TYPE ST_PolarIIChamber_HolderRotateServiceCtrl :
STRUCT
	OPR : ST_ServiceCtrl;
	MoveVelocityCW : ST_ServiceCtrl;
	MoveVelocityCCW : ST_ServiceCtrl;
	MoveModulo : ST_ServiceCtrl;
END_STRUCT
END_TYPE

(* stored: Version 1.1.0.1, ProductVersion 3.1.4026.18
   DUT ST_PolarIIChamber_HolderRotateServiceCtrl: Id {14000000-0000-0000-0000-000000000043} *)
